Fanuc KAREL source: KO00029.KL

PROGRAM KO00029
%NOLOCKGROUP
VAR
  P1: JOINTPOS
  P2: JOINTPOS
  P3: JOINTPOS
  P4: JOINTPOS
  OUT: POSITION
BEGIN
  OUT = FRAME(P1, P2, P3, P4)
END KO00029
